FUNCTION_BLOCK E_MUX_FIFO_2_Adapter (* Adapter-Variante von FIFO::E_MUX_FIFO_2: merkt sich bei EI1/EI2 den Kanal (0/1) in einer FIFO und liefert ihn ueber den Plug OUT_DATA (AFIFO_UINT, Kanal in OUT) einzeln aus. PROCESSED kommt ueber den Rueckkanal. Gegenstueck: E_DEMUX_FIFO_2. *)
  (* Standard: 61499-2; Description: Copyright (c) 2026 Meisterschulen am Ostbahnhof This program and the accompanying materials are made available under the terms of the Eclipse Public License 2.0 which is available at https://www.eclipse.org/legal/epl-2.0/ SPDX-License-Identifier: EPL-2.0 *)
  (* Version 1.0, 2026-11-11, Franz Höpfinger, Meisterschulen am Ostbahnhof, Neu auf Basis von FIFO_UINT_Adapter 1.1: PUSH/IN durch EI1/EI2 ersetzt, der Kanal wird beim Eintreffen des Ereignisses im FB gespeichert und als OUT ueber AFIFO_UINT geliefert. *)
  PACKAGE FIFO_adapter;
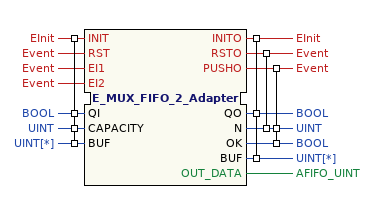
  EVENT_INPUT
    INIT : EInit WITH QI, CAPACITY, BUF; (* Service Initialization *)
    RST; (* Queue leeren und Liefer-Sperre aufheben - Reset der ganzen Kette, der Konsument muss mit zurueckgesetzt werden *)
    EI1; (* Kanal 1 (0) ans Ende der Queue anhaengen, falls Platz vorhanden *)
    EI2; (* Kanal 2 (1) ans Ende der Queue anhaengen, falls Platz vorhanden *)
  END_EVENT
  EVENT_OUTPUT
    INITO : EInit WITH QO, BUF; (* Initialisierung bestaetigt *)
    RSTO WITH N; (* Reset bestaetigt *)
    PUSHO WITH N, OK; (* EI1/EI2 bestaetigt (OK=FALSE wenn Queue voll war oder QO=FALSE) *)
  END_EVENT
  VAR_INPUT
    QI : BOOL; (* Event Input Qualifier *)
    CAPACITY : UINT; (* Kapazitaet - MUSS der Anzahl Elemente von BUF entsprechen, daher immer ueber F_LEN_ARRAY hinter der PROVIDE_ARR_x_UINT-Instanz ermitteln. Ein groesserer Wert schreibt ueber BUF hinaus. 0 ergibt QO=FALSE. *)
  END_VAR
  VAR_OUTPUT
    QO : BOOL; (* Event Output Qualifier *)
    N : UINT; (* Anzahl aktuell wartender (noch nicht ausgelieferter) Elemente *)
    OK : BOOL; (* TRUE wenn das letzte EI1/EI2 erfolgreich war (Queue war nicht voll und QO=TRUE) *)
  END_VAR
  VAR_IN_OUT
    BUF : ARRAY [*] OF UINT; (* Ringpuffer fuer die Kanalnummern --Speicher - Groesse wird extern ueber eine angeschlossene PROVIDE_ARR_x_UINT-Instanz vorgegeben *)
  END_VAR
  PLUGS
    OUT_DATA : FIFO_adapter::AFIFO_UINT; (* Konsument haengt per Socket hier an - DATA liefert den naechsten Wert, PROCESSED (Rueckkanal) quittiert *)
  END_PLUGS
  VAR
    PTR : UINT; (* Schreibposition fuer das naechste EI1/EI2 *)
    KIN : UINT; (* Kanal des gerade eingetroffenen Ereignisses *)
    OUTPTR : UINT; (* Leseposition fuer den naechsten auszuliefernden Wert *)
    DELIVERING : BOOL; (* TRUE = ein Wert wurde per OUT_DATA.DATA geliefert, auf OUT_DATA.PROCESSED wird gewartet *)
  END_VAR
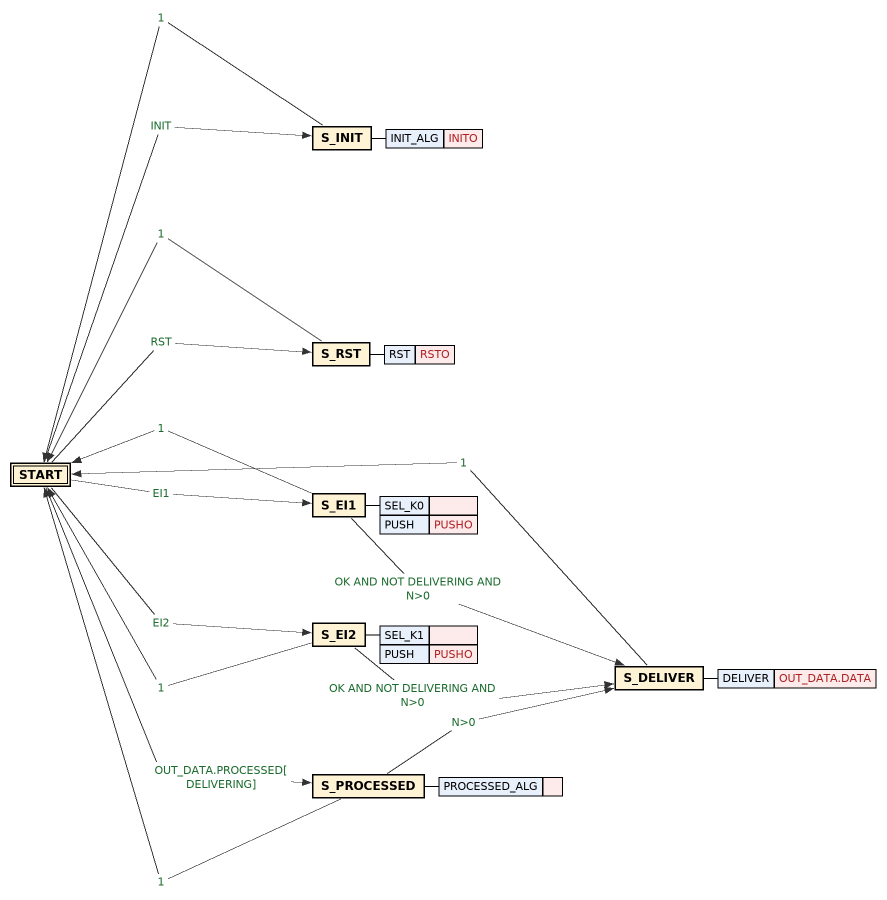
  EC_STATES
    START; (* Initial State *)
    S_INIT : INIT_ALG -> INITO;
    S_RST : RST -> RSTO;
    S_EI1 : SEL_K0, PUSH -> PUSHO;
    S_EI2 : SEL_K1, PUSH -> PUSHO;
    S_PROCESSED : PROCESSED_ALG;
    S_DELIVER : DELIVER -> OUT_DATA.DATA; (* Naechsten Wert aus der Queue entnehmen und ueber den Plug ausliefern *)
  END_STATES
  EC_TRANSITIONS
    START TO S_INIT := INIT;
    START TO S_RST := RST;
    START TO S_EI1 := EI1;
    START TO S_EI2 := EI2;
    START TO S_PROCESSED := OUT_DATA.PROCESSED[DELIVERING];
    S_INIT TO START := 1;
    S_RST TO START := 1;
    S_EI1 TO S_DELIVER := OK AND NOT DELIVERING AND N>0;
    S_EI1 TO START := 1;
    S_EI2 TO S_DELIVER := OK AND NOT DELIVERING AND N>0;
    S_EI2 TO START := 1;
    S_PROCESSED TO S_DELIVER := N>0;
    S_PROCESSED TO START := 1;
    S_DELIVER TO START := 1;
  END_TRANSITIONS
  ALGORITHM INIT_ALG IN ST: (* Queue leeren und QI/QO durchreichen *)
PTR := 0;
OUTPTR := 0;
N := 0;
DELIVERING := FALSE;
OK := FALSE;
QO := QI AND CAPACITY > 0;
  END_ALGORITHM
  ALGORITHM RST IN ST: (* Queue und Liefer-Sperre leeren - RST setzt die ganze Kette zurueck, der Konsument muss mit zurueckgesetzt werden *)
PTR := 0;
OUTPTR := 0;
N := 0;
DELIVERING := FALSE;
OK := FALSE;
  END_ALGORITHM
  ALGORITHM SEL_K0 IN ST: (* Kanal 1 *)
KIN := 0;
  END_ALGORITHM
  ALGORITHM SEL_K1 IN ST: (* Kanal 2 *)
KIN := 1;
  END_ALGORITHM
  ALGORITHM PUSH IN ST: (* Kanal anhaengen, falls Platz vorhanden *)
IF NOT QO OR N >= CAPACITY THEN
    OK := FALSE;
ELSE
    OK := TRUE;
    BUF[PTR] := KIN;
    PTR := (PTR + 1) MOD CAPACITY;
    N := N + 1;
END_IF;
  END_ALGORITHM
  ALGORITHM PROCESSED_ALG IN ST: (* Liefer-Sperre aufheben - das naechste DATA folgt ueber die Transition nach S_DELIVER, falls die Queue noch Elemente enthaelt *)
DELIVERING := FALSE;
  END_ALGORITHM
  ALGORITHM DELIVER IN ST: (* Vordersten Wert entnehmen und ueber den Plug liefern *)
OUT_DATA.OUT := BUF[OUTPTR];
OUTPTR := (OUTPTR + 1) MOD CAPACITY;
N := N - 1;
OUT_DATA.N := N;
DELIVERING := TRUE;
  END_ALGORITHM
END_FUNCTION_BLOCK
